FUNCTION_BLOCK "FB_CraneSpeedCheck"
{ S7_Optimized_Access := 'TRUE' }
VERSION : 0.1
   VAR_INPUT
      LeftSpeed10 : INT;
      RightSpeed10 : INT;
      ReferenceSpeed10 : INT;
   END_VAR
   VAR_OUTPUT
      SyncOK : BOOL;
      SyncBad : BOOL;
      Invalid : BOOL;
   END_VAR
   VAR_TEMP
      tmpValid : BOOL;
      tmpLeft : DINT;
      tmpRight : DINT;
      tmpRef : DINT;
      tmpDiff12 : DINT;
      tmpSumRatio : DINT;
      tmpRatioTarget : DINT;
      tmpSyncCond : BOOL;
      tmpRatioCond : BOOL;
   END_VAR
BEGIN

      // 每周期先复位所有输出，保证恰好一个为 TRUE
      #SyncOK := FALSE;
      #SyncBad := FALSE;
      #Invalid := FALSE;

      // 拓宽为 DINT 后再进行后续运算，避免 INT 溢出
      #tmpLeft := INT_TO_DINT(#LeftSpeed10);
      #tmpRight := INT_TO_DINT(#RightSpeed10);
      #tmpRef := INT_TO_DINT(#ReferenceSpeed10);

      // 量程校验：三路均在 0..100，且参考速度 > 0
      #tmpValid := (#tmpLeft >= 0) AND (#tmpLeft <= 100)
                   AND (#tmpRight >= 0) AND (#tmpRight <= 100)
                   AND (#tmpRef > 0) AND (#tmpRef <= 100);

      IF NOT #tmpValid THEN
         #Invalid := TRUE;
      ELSE
         // 同步约束：|L - R| <= 1
         #tmpDiff12 := #tmpLeft - #tmpRight;
         IF #tmpDiff12 < 0 THEN
            #tmpDiff12 := -#tmpDiff12;
         END_IF;
         #tmpSyncCond := (#tmpDiff12 <= 1);

         // 传动比约束：|L + R - 13 * Ref| <= 2
         #tmpRatioTarget := 13 * #tmpRef;
         #tmpSumRatio := #tmpLeft + #tmpRight - #tmpRatioTarget;
         IF #tmpSumRatio < 0 THEN
            #tmpSumRatio := -#tmpSumRatio;
         END_IF;
         #tmpRatioCond := (#tmpSumRatio <= 2);

         IF #tmpSyncCond AND #tmpRatioCond THEN
            #SyncOK := TRUE;
         ELSE
            #SyncBad := TRUE;
         END_IF;
      END_IF;

END_FUNCTION_BLOCK